Staubli VAL3: MatrixLib.dtx


